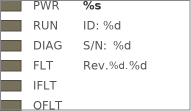
VISUALIZATION FRM_ModuleStatus  // 191x111
VAR_IN_OUT
    bPower: BOOL;
    bRun: BOOL;
    bDiag: BOOL;
    bFault: BOOL;
    bInputFault: BOOL;
    bOutputFault: BOOL;
    sName: STRING;
    nID: UDINT;
    nSerialNumber: UDINT;
   anRevision: ARRAY [1..2] OF BYTE;
END_VAR
    Rectangle (0,0 21x11), colour toggle: bPower
    Rectangle (0,20 21x11), colour toggle: bRun
    Rectangle (0,40 21x11), colour toggle: bDiag
    Rectangle (0,60 21x11), colour toggle: bFault
    Rectangle (0,80 21x11), colour toggle: bInputFault
    Rectangle (0,100 21x11), colour toggle: bOutputFault
    Label (30,0 41x11), "PWR"
    Label (30,20 41x11), "RUN"
    Label (30,40 41x11), "DIAG"
    Label (30,60 41x11), "FLT"
    Label (30,80 41x11), "IFLT"
    Label (30,100 41x11), "OFLT"
    Textfield (110,40 81x11), "%d", text variable: nSerialNumber
    Textfield (100,20 91x11), "%d", text variable: nID
    Textfield (80,0 111x11), "%s", text variable: sName
    Label (80,20 21x11), "ID:"
    Label (80,40 31x11), "S/N:"
    Textfield (110,60 21x11), "%d.", text variable: anRevision[1]
    Label (80,60 31x11), "Rev."
    Textfield (126,60 21x11), "%d", text variable: anRevision[2]
END_VISUALIZATION

(* stored: Version 1.1.0.1
   Visu FRM_ModuleStatus: Id {58c5cd6b-1cf3-04aa-3c8a-12fb61bd275d} *)
